Fanuc KAREL source: kd00002.KL

-- PROVISIONAL review KL for V770-1; original PC SHA256 ee8df7a8b48bf6f5dfad081f141001b7cad62b20ede5734c5b572f6b56b10f98
-- Incomplete behavior may be omitted. Consult companion uncertainty JSON. Do not deploy.
PROGRAM KD00002
%NOLOCKGROUP
VAR
  I : INTEGER
  J : INTEGER
  B : BOOLEAN
  R : REAL
  S : STRING[80]
BEGIN
  -- UNRESOLVED_PC offsets 5-12; opcodes 9D,23
  -- UNRESOLVED_PC offsets 17-21; opcodes 7F
END KD00002
